// TIA Portal V20 export
DATA_BLOCK "DB_LASER"   // DB402
{ S7_Optimized_Access := 'TRUE' }
// stored: AutoNumber false, MemoryReserve 100
   VAR
      DATA_DO_ETIKETY : Struct
         TEXT : String[5];
         "INT" : Int;
         "REAL" : Real;
         PROGRAM : Array[0..1] of String[10];
      END_STRUCT;
      DATA_DO_DAT : Struct
         ZAVORKA_L : Char := '<';
         ZAVORKA_P : Char := '>';
         XLP : Array[0..3] of Char;
      END_STRUCT;
      smaz_me_start : Bool;
      smaz_me_adresa : Int;
   END_VAR
BEGIN
   DATA_DO_ETIKETY.PROGRAM[0] := 'TEST_1';
   DATA_DO_ETIKETY.PROGRAM[1] := 'TEST_222';
   DATA_DO_DAT.XLP[0] := '.';
   DATA_DO_DAT.XLP[1] := 'x';
   DATA_DO_DAT.XLP[2] := 'l';
   DATA_DO_DAT.XLP[3] := 'p';
END_DATA_BLOCK
